Fanuc KAREL source: kb00037.KL

-- PROVISIONAL review KL for V1013-1; original PC SHA256 a150f1b14411422f27935e572728f4d9fb2910d53577489afa08c9331ca63e04
-- Incomplete behavior may be omitted. Consult companion uncertainty JSON. Do not deploy.
PROGRAM KB00037
%NOLOCKGROUP
BEGIN
  -- UNRESOLVED_PC offsets 5-16; opcodes 2E,23
  -- UNRESOLVED_PC offsets 21-28; opcodes 9D,23
  -- UNRESOLVED_PC offsets 33-40; opcodes 9D,23
  -- UNRESOLVED_PC offsets 45-54; opcodes 3F,75
  -- UNRESOLVED_PC offsets 59-89; opcodes 27,22,22,22,22,2A,31
  -- UNRESOLVED_PC offsets 94-98; opcodes 7F
END KB00037
